SUBAPPLICATION Station_Alive_VT_OPC (* Verbindungsueberwachung einer Station ueber ihren Tick: Status-Button gruen/rot, Abbrueche und Boots auf dem VT *)
  (* Standard: 61499-2; Description: Copyright (c) 2026 Meisterschulen am Ostbahnhof This program and the accompanying materials are made available under the terms of the Eclipse Public License 2.0 which is available at https://www.eclipse.org/legal/epl-2.0/ SPDX-License-Identifier: EPL-2.0 *)
  (* Version 1.0, 2026-10-29, Franz Höpfinger, Meisterschulen am Ostbahnhof, Neu: Tick der Station (SystemTickSender_OPC, 200 ms) per Remote-Subscribe, E_RDELAY als Timeout. ALIVE geht beim ersten Tick auf TRUE, nach DT ohne Tick auf FALSE. Jede fallende Flanke zaehlt als Abbruch, BOOT-Ereignisse (von Boot_Zaehler_OPC) als Boots. *)
  PACKAGE MyLib::sys;
  IMPORT isobus::UT::Q::const::IDs::ID_NULL;
  (* Documentation:
  Verbindungsüberwachung einer Station
   Jede Station veröffentlicht alle 200 ms ihren Tick (SystemTickSender_OPC). Dieser Baustein abonniert ihn auf STG1. Jeder Tick setzt ALIVE und startet den Timeout DT neu. Kommt DT lang kein Tick, fällt ALIVE auf FALSE.
    - Status-Button: grün bei ALIVE, rot sonst (Pool-Startwert rot, bis der erste Tick kommt).
   - Abbrüche: jede fallende Flanke von ALIVE.
   - Boots: jedes Ereignis an BOOT (von Boot_Zaehler_OPC).
    Beide Zähler laufen im RAM und beginnen beim Start von STG1 bei 0.
  *)
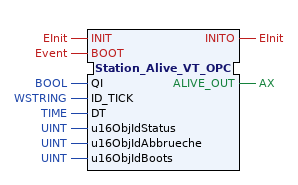
  EVENT_INPUT
    INIT : EInit; (* Initialization Request *)
    BOOT; (* Station hat ihren Start gemeldet *)
  END_EVENT
  EVENT_OUTPUT
    INITO : EInit; (* Initialization Confirm *)
  END_EVENT
  VAR_INPUT
    QI : BOOL := TRUE; (* Quality Input - TRUE to enable service *)
    ID_TICK : WSTRING; (* Remote-Subscribe auf den Tick der Station *)
    DT : TIME := T#2s; (* Timeout ohne Tick *)
    u16ObjIdStatus : UINT := ID_NULL; (* Status-Button (gruen/rot) *)
    u16ObjIdAbbrueche : UINT := ID_NULL; (* NumberVariable Abbrueche *)
    u16ObjIdBoots : UINT := ID_NULL; (* NumberVariable Boots *)
  END_VAR
  PLUGS
    ALIVE_OUT : adapter::types::unidirectional::AX; (* TRUE solange Ticks kommen *)
  END_PLUGS
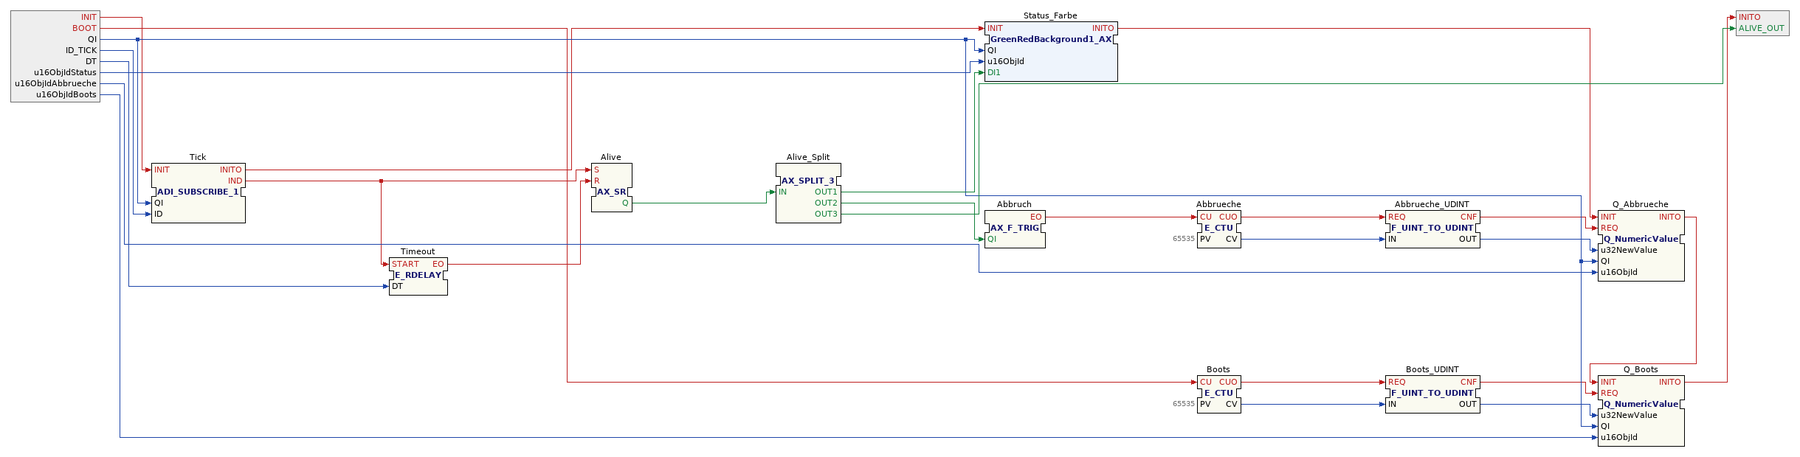
  FBS
    Tick : adapter::net::ADI_SUBSCRIBE_1;
    Timeout : iec61499::events::E_RDELAY;
    Alive : adapter::events::unidirectional::AX_SR;
    Alive_Split : adapter::events::unidirectional::AX_SPLIT_3;
    Abbruch : adapter::events::unidirectional::AX_F_TRIG;
    Abbrueche : iec61499::events::E_CTU(PV := 65535);
    Abbrueche_UDINT : iec61131::conversion::F_UINT_TO_UDINT;
    Q_Abbrueche : isobus::UT::Q::Q_NumericValue;
    Boots : iec61499::events::E_CTU(PV := 65535);
    Boots_UDINT : iec61131::conversion::F_UINT_TO_UDINT;
    Q_Boots : isobus::UT::Q::Q_NumericValue;
  END_FBS
  SUBAPPS
    Status_Farbe : MyLib::sys::GreenRedBackground1_AX;
  END_SUBAPPS
  EVENT_CONNECTIONS
    INIT TO Tick.INIT;
    Tick.INITO TO Status_Farbe.INIT;
    Status_Farbe.INITO TO Q_Abbrueche.INIT;
    Q_Abbrueche.INITO TO Q_Boots.INIT;
    Q_Boots.INITO TO INITO;
    Tick.IND TO Timeout.START;
    Tick.IND TO Alive.S;
    Timeout.EO TO Alive.R;
    Abbruch.EO TO Abbrueche.CU;
    Abbrueche.CUO TO Abbrueche_UDINT.REQ;
    Abbrueche_UDINT.CNF TO Q_Abbrueche.REQ;
    BOOT TO Boots.CU;
    Boots.CUO TO Boots_UDINT.REQ;
    Boots_UDINT.CNF TO Q_Boots.REQ;
  END_CONNECTIONS
  DATA_CONNECTIONS
    QI TO Tick.QI;
    ID_TICK TO Tick.ID;
    DT TO Timeout.DT;
    QI TO Status_Farbe.QI;
    u16ObjIdStatus TO Status_Farbe.u16ObjId;
    Abbrueche.CV TO Abbrueche_UDINT.IN;
    Abbrueche_UDINT.OUT TO Q_Abbrueche.u32NewValue;
    QI TO Q_Abbrueche.QI;
    u16ObjIdAbbrueche TO Q_Abbrueche.u16ObjId;
    Boots.CV TO Boots_UDINT.IN;
    Boots_UDINT.OUT TO Q_Boots.u32NewValue;
    QI TO Q_Boots.QI;
    u16ObjIdBoots TO Q_Boots.u16ObjId;
  END_CONNECTIONS
  ADAPTER_CONNECTIONS
    Alive.Q TO Alive_Split.IN;
    Alive_Split.OUT1 TO Status_Farbe.DI1;
    Alive_Split.OUT2 TO Abbruch.QI;
    Alive_Split.OUT3 TO ALIVE_OUT;
  END_CONNECTIONS
END_SUBAPPLICATION
